Fanuc KAREL source: KT00542.KL

PROGRAM KT00542
%NOLOCKGROUP
VAR
  P1: JOINTPOS
  P2: XYZWPR
  OUT: JOINTPOS
BEGIN
    P2.Y = 2.0
  OUT = P1 : P2
END KT00542
